(* PLC project Vn_fbd_neg_output, Beckhoff Automation GmbH TwinCAT PLC Control 3.5.13.21 *)
(* stored: creationDateTime 1970-01-01T00:00:00 *)

PROGRAM Vn_fbd_neg_output

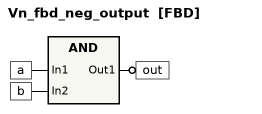
(* FBD diagram, written out as Structured Text *)
out := NOT (a AND b);
END_PROGRAM
